Fanuc KAREL source: KB00042.KL

PROGRAM KB00042
%NOLOCKGROUP
%ENVIRONMENT TIM
VAR
  P1: STRING[80]
  P2: INTEGER
BEGIN
  P1 = 'A'
  P2 = 1
  CNV_STR_TIME(P1, P2)
END KB00042
